(* IEC 61131-3 sources: llm-plc-st-eval/data/processed_definitivo/gemini-3.1-pro-preview/B2/few_shot, 3 files *)

(* ---- ejec_1.st ---- *)
FUNCTION_BLOCK FB_Valvula
VAR_INPUT
    nivelAlto : BOOL; (* Sensor de nivel alto *)
END_VAR
VAR_OUTPUT
    valvula : BOOL; (* Valvula de drenaje *)
END_VAR
VAR
    tRetardo : TON; (* Temporizador de retardo a la conexion *)
END_VAR

(* La valvula abre tras 5 s continuos de nivel alto y cierra de inmediato si baja *)
tRetardo(IN := nivelAlto, PT := T#5S);
valvula := tRetardo.Q;
END_FUNCTION_BLOCK

(* ---- ejec_2.st ---- *)
FUNCTION_BLOCK FB_Valvula
VAR_INPUT
    nivelAlto : BOOL; (* Sensor de nivel alto *)
END_VAR
VAR_OUTPUT
    valvula : BOOL; (* Valvula de drenaje *)
END_VAR
VAR
    tRetardo : TON; (* Temporizador de retardo a la conexion *)
END_VAR

(* Retardo de 5 s para abrir la valvula; cierra de inmediato al desactivarse el sensor *)
tRetardo(IN := nivelAlto, PT := T#5S);
valvula := tRetardo.Q;
END_FUNCTION_BLOCK

(* ---- ejec_3.st ---- *)
FUNCTION_BLOCK FB_Valvula
VAR_INPUT
    nivelAlto : BOOL; (* Sensor de nivel alto *)
END_VAR
VAR_OUTPUT
    valvula : BOOL; (* Valvula de drenaje *)
END_VAR
VAR
    tRetardo : TON; (* Temporizador de retardo a la conexion *)
END_VAR

(* Retardo de 5 s para abrir la valvula; cierre inmediato al desactivarse el sensor *)
tRetardo(IN := nivelAlto, PT := T#5S);
valvula := tRetardo.Q;
END_FUNCTION_BLOCK
